Yaskawa INFORM job: PAT_POSTYPE_PULSE.JBI

/JOB
//NAME PAT_POSTYPE_PULSE
//POS
///NPOS 7,0,0,0,0,0
///TOOL 0
///POSTYPE PULSE
///PULSE
C00000=1200,-35000,21000,0,-48000,500
C00001=1200,-41000,9000,0,-52000,500
C00002=1200,-38000,15000,0,-50000,500
C00003=-9800,-38000,15000,0,-50000,-9200
C00004=-9800,-42000,7000,0,-53000,-9200
C00005=-9800,-38000,15000,0,-50000,-9200
C00006=1200,-35000,21000,0,-48000,500
//INST
///DATE 2026/11/02 14:40
///ATTR SC,RW
///GROUP1 RB1
NOP
'SYNTHETIC TEST DATA - NOT A REAL ROBOT JOB
MOVL C00000 V=200.0
MOVL C00001 V=80.0
DOUT OT#(1) ON
TIMER T=0.50
MOVL C00002 V=80.0
MOVL C00003 V=250.0
MOVL C00004 V=80.0
TIMER T=3.00
DOUT OT#(1) OFF
TIMER T=0.50
MOVL C00005 V=80.0
MOVL C00006 V=200.0
END
